FUNCTION_BLOCK PID_GAIN_TRANSITION (* Experimental; offline checks only; native export/runtime pending *)
  (* Standard: 61499-2 *)
  (* Version 0.1, 2026-10-20, Guilherme *)
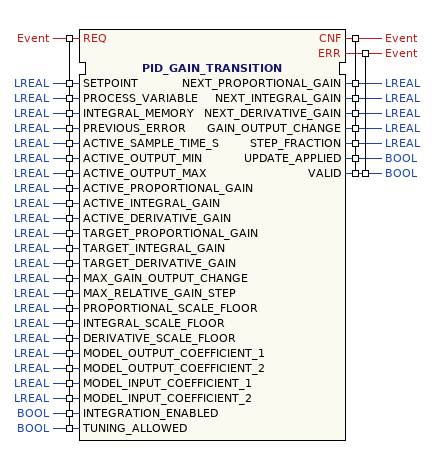
  EVENT_INPUT
    REQ WITH SETPOINT, PROCESS_VARIABLE, INTEGRAL_MEMORY, PREVIOUS_ERROR, ACTIVE_SAMPLE_TIME_S, ACTIVE_OUTPUT_MIN, ACTIVE_OUTPUT_MAX, ACTIVE_PROPORTIONAL_GAIN, ACTIVE_INTEGRAL_GAIN, ACTIVE_DERIVATIVE_GAIN, TARGET_PROPORTIONAL_GAIN, TARGET_INTEGRAL_GAIN, TARGET_DERIVATIVE_GAIN, MAX_GAIN_OUTPUT_CHANGE, MAX_RELATIVE_GAIN_STEP, PROPORTIONAL_SCALE_FLOOR, INTEGRAL_SCALE_FLOOR, DERIVATIVE_SCALE_FLOOR, MODEL_OUTPUT_COEFFICIENT_1, MODEL_OUTPUT_COEFFICIENT_2, MODEL_INPUT_COEFFICIENT_1, MODEL_INPUT_COEFFICIENT_2, INTEGRATION_ENABLED, TUNING_ALLOWED;
  END_EVENT
  EVENT_OUTPUT
    CNF WITH NEXT_PROPORTIONAL_GAIN, NEXT_INTEGRAL_GAIN, NEXT_DERIVATIVE_GAIN, GAIN_OUTPUT_CHANGE, STEP_FRACTION, UPDATE_APPLIED, VALID;
    ERR WITH VALID;
  END_EVENT
  VAR_INPUT
    SETPOINT : LREAL;
    PROCESS_VARIABLE : LREAL;
    INTEGRAL_MEMORY : LREAL;
    PREVIOUS_ERROR : LREAL;
    ACTIVE_SAMPLE_TIME_S : LREAL;
    ACTIVE_OUTPUT_MIN : LREAL;
    ACTIVE_OUTPUT_MAX : LREAL;
    ACTIVE_PROPORTIONAL_GAIN : LREAL;
    ACTIVE_INTEGRAL_GAIN : LREAL;
    ACTIVE_DERIVATIVE_GAIN : LREAL;
    TARGET_PROPORTIONAL_GAIN : LREAL;
    TARGET_INTEGRAL_GAIN : LREAL;
    TARGET_DERIVATIVE_GAIN : LREAL;
    MAX_GAIN_OUTPUT_CHANGE : LREAL;
    MAX_RELATIVE_GAIN_STEP : LREAL;
    PROPORTIONAL_SCALE_FLOOR : LREAL;
    INTEGRAL_SCALE_FLOOR : LREAL;
    DERIVATIVE_SCALE_FLOOR : LREAL;
    MODEL_OUTPUT_COEFFICIENT_1 : LREAL;
    MODEL_OUTPUT_COEFFICIENT_2 : LREAL;
    MODEL_INPUT_COEFFICIENT_1 : LREAL;
    MODEL_INPUT_COEFFICIENT_2 : LREAL;
    INTEGRATION_ENABLED : BOOL;
    TUNING_ALLOWED : BOOL;
  END_VAR
  VAR_OUTPUT
    NEXT_PROPORTIONAL_GAIN : LREAL;
    NEXT_INTEGRAL_GAIN : LREAL;
    NEXT_DERIVATIVE_GAIN : LREAL;
    GAIN_OUTPUT_CHANGE : LREAL;
    STEP_FRACTION : LREAL;
    UPDATE_APPLIED : BOOL;
    VALID : BOOL;
  END_VAR
  VAR
    CURRENT_ERROR : LREAL;
    NEXT_INTEGRAL : LREAL;
    CURRENT_DERIVATIVE : LREAL;
    OLD_RAW : LREAL;
    NEW_RAW : LREAL;
    DELTA_P : LREAL;
    DELTA_I : LREAL;
    DELTA_D : LREAL;
    FULL_EFFECT : LREAL;
    MAGNITUDE : LREAL;
    SCALE : LREAL;
    RELATIVE_STEP : LREAL;
    FRACTION_LIMIT : LREAL;
    CANDIDATE_P : LREAL;
    CANDIDATE_I : LREAL;
    CANDIDATE_D : LREAL;
    Q0 : LREAL;
    Q1 : LREAL;
    Q2 : LREAL;
    A1 : LREAL;
    A2 : LREAL;
    A3 : LREAL;
    A4 : LREAL;
    DENOMINATOR : LREAL;
    B1 : LREAL;
    B2 : LREAL;
    B3 : LREAL;
    C1 : LREAL;
    C2 : LREAL;
    D1 : LREAL;
    CANDIDATE_VALID : BOOL;
  END_VAR
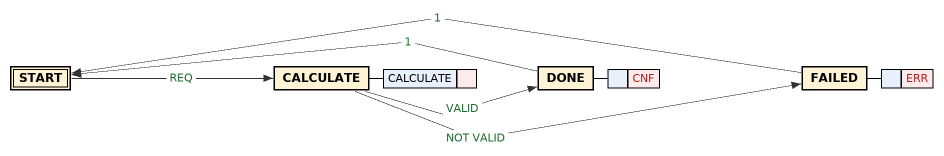
  EC_STATES
    START;
    CALCULATE : CALCULATE;
    DONE : -> CNF;
    FAILED : -> ERR;
  END_STATES
  EC_TRANSITIONS
    START TO CALCULATE := REQ;
    CALCULATE TO DONE := VALID;
    CALCULATE TO FAILED := NOT VALID;
    DONE TO START := 1;
    FAILED TO START := 1;
  END_TRANSITIONS
  ALGORITHM CALCULATE IN ST:
VALID := (SETPOINT >= -1.0E+100) AND (SETPOINT <= 1.0E+100) AND (PROCESS_VARIABLE >= -1.0E+100) AND (PROCESS_VARIABLE <= 1.0E+100) AND (INTEGRAL_MEMORY >= -1.0E+100) AND (INTEGRAL_MEMORY <= 1.0E+100) AND (PREVIOUS_ERROR >= -1.0E+100) AND (PREVIOUS_ERROR <= 1.0E+100) AND (ACTIVE_SAMPLE_TIME_S >= -1.0E+100) AND (ACTIVE_SAMPLE_TIME_S <= 1.0E+100) AND (ACTIVE_OUTPUT_MIN >= -1.0E+100) AND (ACTIVE_OUTPUT_MIN <= 1.0E+100) AND (ACTIVE_OUTPUT_MAX >= -1.0E+100) AND (ACTIVE_OUTPUT_MAX <= 1.0E+100) AND (ACTIVE_PROPORTIONAL_GAIN >= -1.0E+100) AND (ACTIVE_PROPORTIONAL_GAIN <= 1.0E+100) AND (ACTIVE_INTEGRAL_GAIN >= -1.0E+100) AND (ACTIVE_INTEGRAL_GAIN <= 1.0E+100) AND (ACTIVE_DERIVATIVE_GAIN >= -1.0E+100) AND (ACTIVE_DERIVATIVE_GAIN <= 1.0E+100) AND (MAX_GAIN_OUTPUT_CHANGE >= -1.0E+100) AND (MAX_GAIN_OUTPUT_CHANGE <= 1.0E+100) AND (MAX_RELATIVE_GAIN_STEP >= -1.0E+100) AND (MAX_RELATIVE_GAIN_STEP <= 1.0E+100) AND (PROPORTIONAL_SCALE_FLOOR >= -1.0E+100) AND (PROPORTIONAL_SCALE_FLOOR <= 1.0E+100) AND (INTEGRAL_SCALE_FLOOR >= -1.0E+100) AND (INTEGRAL_SCALE_FLOOR <= 1.0E+100) AND (DERIVATIVE_SCALE_FLOOR >= -1.0E+100) AND (DERIVATIVE_SCALE_FLOOR <= 1.0E+100) AND (ACTIVE_SAMPLE_TIME_S > 0.0) AND (ACTIVE_OUTPUT_MIN < ACTIVE_OUTPUT_MAX) AND (MAX_GAIN_OUTPUT_CHANGE > 0.0) AND (MAX_RELATIVE_GAIN_STEP > 0.0) AND (MAX_RELATIVE_GAIN_STEP <= 1.0) AND (PROPORTIONAL_SCALE_FLOOR > 0.0) AND (INTEGRAL_SCALE_FLOOR > 0.0) AND (DERIVATIVE_SCALE_FLOOR > 0.0);
UPDATE_APPLIED := FALSE;
GAIN_OUTPUT_CHANGE := 0.0;
STEP_FRACTION := 0.0;
IF VALID THEN
NEXT_PROPORTIONAL_GAIN := ACTIVE_PROPORTIONAL_GAIN;
NEXT_INTEGRAL_GAIN := ACTIVE_INTEGRAL_GAIN;
NEXT_DERIVATIVE_GAIN := ACTIVE_DERIVATIVE_GAIN;
IF TUNING_ALLOWED AND INTEGRATION_ENABLED THEN
CANDIDATE_VALID := (TARGET_PROPORTIONAL_GAIN >= -1.0E+100) AND (TARGET_PROPORTIONAL_GAIN <= 1.0E+100) AND (TARGET_INTEGRAL_GAIN >= -1.0E+100) AND (TARGET_INTEGRAL_GAIN <= 1.0E+100) AND (TARGET_DERIVATIVE_GAIN >= -1.0E+100) AND (TARGET_DERIVATIVE_GAIN <= 1.0E+100) AND (MODEL_OUTPUT_COEFFICIENT_1 >= -1.0E+100) AND (MODEL_OUTPUT_COEFFICIENT_1 <= 1.0E+100) AND (MODEL_OUTPUT_COEFFICIENT_2 >= -1.0E+100) AND (MODEL_OUTPUT_COEFFICIENT_2 <= 1.0E+100) AND (MODEL_INPUT_COEFFICIENT_1 >= -1.0E+100) AND (MODEL_INPUT_COEFFICIENT_1 <= 1.0E+100) AND (MODEL_INPUT_COEFFICIENT_2 >= -1.0E+100) AND (MODEL_INPUT_COEFFICIENT_2 <= 1.0E+100) AND (TARGET_PROPORTIONAL_GAIN >= 0.0) AND (TARGET_INTEGRAL_GAIN >= 0.0) AND (TARGET_DERIVATIVE_GAIN >= 0.0);
IF CANDIDATE_VALID THEN
CURRENT_ERROR := SETPOINT - PROCESS_VARIABLE;
NEXT_INTEGRAL := INTEGRAL_MEMORY + ACTIVE_SAMPLE_TIME_S / 2.0 * (CURRENT_ERROR + PREVIOUS_ERROR);
CURRENT_DERIVATIVE := (CURRENT_ERROR - PREVIOUS_ERROR) / ACTIVE_SAMPLE_TIME_S;
OLD_RAW := ACTIVE_PROPORTIONAL_GAIN * CURRENT_ERROR + ACTIVE_INTEGRAL_GAIN * NEXT_INTEGRAL + ACTIVE_DERIVATIVE_GAIN * CURRENT_DERIVATIVE;
DELTA_P := TARGET_PROPORTIONAL_GAIN - ACTIVE_PROPORTIONAL_GAIN;
DELTA_I := TARGET_INTEGRAL_GAIN - ACTIVE_INTEGRAL_GAIN;
DELTA_D := TARGET_DERIVATIVE_GAIN - ACTIVE_DERIVATIVE_GAIN;
FULL_EFFECT := DELTA_P * CURRENT_ERROR + DELTA_I * NEXT_INTEGRAL + DELTA_D * CURRENT_DERIVATIVE;
CANDIDATE_VALID := (CURRENT_ERROR >= -1.0E+100) AND (CURRENT_ERROR <= 1.0E+100) AND (NEXT_INTEGRAL >= -1.0E+100) AND (NEXT_INTEGRAL <= 1.0E+100) AND (CURRENT_DERIVATIVE >= -1.0E+100) AND (CURRENT_DERIVATIVE <= 1.0E+100) AND (OLD_RAW >= -1.0E+100) AND (OLD_RAW <= 1.0E+100) AND (FULL_EFFECT >= -1.0E+100) AND (FULL_EFFECT <= 1.0E+100) AND (OLD_RAW >= ACTIVE_OUTPUT_MIN) AND (OLD_RAW <= ACTIVE_OUTPUT_MAX);
IF CANDIDATE_VALID THEN
STEP_FRACTION := 1.0;
MAGNITUDE := FULL_EFFECT;
IF MAGNITUDE < 0.0 THEN
MAGNITUDE := -MAGNITUDE;
END_IF;
IF MAGNITUDE > MAX_GAIN_OUTPUT_CHANGE THEN
STEP_FRACTION := MAX_GAIN_OUTPUT_CHANGE / MAGNITUDE;
END_IF;
SCALE := ACTIVE_PROPORTIONAL_GAIN;
IF SCALE < 0.0 THEN
SCALE := -SCALE;
END_IF;
IF SCALE < PROPORTIONAL_SCALE_FLOOR THEN
SCALE := PROPORTIONAL_SCALE_FLOOR;
END_IF;
MAGNITUDE := DELTA_P;
IF MAGNITUDE < 0.0 THEN
MAGNITUDE := -MAGNITUDE;
END_IF;
RELATIVE_STEP := MAGNITUDE / SCALE;
IF RELATIVE_STEP > MAX_RELATIVE_GAIN_STEP THEN
FRACTION_LIMIT := MAX_RELATIVE_GAIN_STEP / RELATIVE_STEP;
IF FRACTION_LIMIT < STEP_FRACTION THEN
STEP_FRACTION := FRACTION_LIMIT;
END_IF;
END_IF;
CANDIDATE_P := ACTIVE_PROPORTIONAL_GAIN + STEP_FRACTION * DELTA_P;
SCALE := ACTIVE_INTEGRAL_GAIN;
IF SCALE < 0.0 THEN
SCALE := -SCALE;
END_IF;
IF SCALE < INTEGRAL_SCALE_FLOOR THEN
SCALE := INTEGRAL_SCALE_FLOOR;
END_IF;
MAGNITUDE := DELTA_I;
IF MAGNITUDE < 0.0 THEN
MAGNITUDE := -MAGNITUDE;
END_IF;
RELATIVE_STEP := MAGNITUDE / SCALE;
IF RELATIVE_STEP > MAX_RELATIVE_GAIN_STEP THEN
FRACTION_LIMIT := MAX_RELATIVE_GAIN_STEP / RELATIVE_STEP;
IF FRACTION_LIMIT < STEP_FRACTION THEN
STEP_FRACTION := FRACTION_LIMIT;
END_IF;
END_IF;
CANDIDATE_I := ACTIVE_INTEGRAL_GAIN + STEP_FRACTION * DELTA_I;
SCALE := ACTIVE_DERIVATIVE_GAIN;
IF SCALE < 0.0 THEN
SCALE := -SCALE;
END_IF;
IF SCALE < DERIVATIVE_SCALE_FLOOR THEN
SCALE := DERIVATIVE_SCALE_FLOOR;
END_IF;
MAGNITUDE := DELTA_D;
IF MAGNITUDE < 0.0 THEN
MAGNITUDE := -MAGNITUDE;
END_IF;
RELATIVE_STEP := MAGNITUDE / SCALE;
IF RELATIVE_STEP > MAX_RELATIVE_GAIN_STEP THEN
FRACTION_LIMIT := MAX_RELATIVE_GAIN_STEP / RELATIVE_STEP;
IF FRACTION_LIMIT < STEP_FRACTION THEN
STEP_FRACTION := FRACTION_LIMIT;
END_IF;
END_IF;
CANDIDATE_D := ACTIVE_DERIVATIVE_GAIN + STEP_FRACTION * DELTA_D;
CANDIDATE_P := ACTIVE_PROPORTIONAL_GAIN + STEP_FRACTION * DELTA_P;
CANDIDATE_I := ACTIVE_INTEGRAL_GAIN + STEP_FRACTION * DELTA_I;
CANDIDATE_D := ACTIVE_DERIVATIVE_GAIN + STEP_FRACTION * DELTA_D;
NEW_RAW := CANDIDATE_P * CURRENT_ERROR + CANDIDATE_I * NEXT_INTEGRAL + CANDIDATE_D * CURRENT_DERIVATIVE;
Q0 := CANDIDATE_P + CANDIDATE_I * ACTIVE_SAMPLE_TIME_S / 2.0 + CANDIDATE_D / ACTIVE_SAMPLE_TIME_S;
Q1 := -CANDIDATE_P + CANDIDATE_I * ACTIVE_SAMPLE_TIME_S / 2.0 - 2.0 * CANDIDATE_D / ACTIVE_SAMPLE_TIME_S;
Q2 := CANDIDATE_D / ACTIVE_SAMPLE_TIME_S;
A1 := -1.0 - MODEL_OUTPUT_COEFFICIENT_1 + MODEL_INPUT_COEFFICIENT_1 * Q0;
A2 := MODEL_OUTPUT_COEFFICIENT_1 - MODEL_OUTPUT_COEFFICIENT_2 + MODEL_INPUT_COEFFICIENT_1 * Q1 + MODEL_INPUT_COEFFICIENT_2 * Q0;
A3 := MODEL_OUTPUT_COEFFICIENT_2 + MODEL_INPUT_COEFFICIENT_1 * Q2 + MODEL_INPUT_COEFFICIENT_2 * Q1;
A4 := MODEL_INPUT_COEFFICIENT_2 * Q2;
CANDIDATE_VALID := (CANDIDATE_P >= -1.0E+100) AND (CANDIDATE_P <= 1.0E+100) AND (CANDIDATE_I >= -1.0E+100) AND (CANDIDATE_I <= 1.0E+100) AND (CANDIDATE_D >= -1.0E+100) AND (CANDIDATE_D <= 1.0E+100) AND (NEW_RAW >= -1.0E+100) AND (NEW_RAW <= 1.0E+100) AND (A1 >= -1.0E+100) AND (A1 <= 1.0E+100) AND (A2 >= -1.0E+100) AND (A2 <= 1.0E+100) AND (A3 >= -1.0E+100) AND (A3 <= 1.0E+100) AND (A4 >= -1.0E+100) AND (A4 <= 1.0E+100) AND (NEW_RAW >= ACTIVE_OUTPUT_MIN) AND (NEW_RAW <= ACTIVE_OUTPUT_MAX);
IF CANDIDATE_VALID THEN
CANDIDATE_VALID := (A4 > -1.0) AND (A4 < 1.0);
IF CANDIDATE_VALID THEN
DENOMINATOR := 1.0 - A4 * A4;
CANDIDATE_VALID := DENOMINATOR > 1.0E-12;
IF CANDIDATE_VALID THEN
B1 := (A1 - A4 * A3) / DENOMINATOR;
B2 := (A2 - A4 * A2) / DENOMINATOR;
B3 := (A3 - A4 * A1) / DENOMINATOR;
CANDIDATE_VALID := (B1 >= -1.0E+100) AND (B1 <= 1.0E+100) AND (B2 >= -1.0E+100) AND (B2 <= 1.0E+100) AND (B3 >= -1.0E+100) AND (B3 <= 1.0E+100);
END_IF;
END_IF;
END_IF;
IF CANDIDATE_VALID THEN
CANDIDATE_VALID := (B3 > -1.0) AND (B3 < 1.0);
IF CANDIDATE_VALID THEN
DENOMINATOR := 1.0 - B3 * B3;
CANDIDATE_VALID := DENOMINATOR > 1.0E-12;
IF CANDIDATE_VALID THEN
C1 := (B1 - B3 * B2) / DENOMINATOR;
C2 := (B2 - B3 * B1) / DENOMINATOR;
CANDIDATE_VALID := (C1 >= -1.0E+100) AND (C1 <= 1.0E+100) AND (C2 >= -1.0E+100) AND (C2 <= 1.0E+100);
END_IF;
END_IF;
END_IF;
IF CANDIDATE_VALID THEN
CANDIDATE_VALID := (C2 > -1.0) AND (C2 < 1.0);
IF CANDIDATE_VALID THEN
DENOMINATOR := 1.0 - C2 * C2;
CANDIDATE_VALID := DENOMINATOR > 1.0E-12;
IF CANDIDATE_VALID THEN
D1 := (C1 - C2 * C1) / DENOMINATOR;
CANDIDATE_VALID := (D1 >= -1.0E+100) AND (D1 <= 1.0E+100);
END_IF;
END_IF;
END_IF;
IF CANDIDATE_VALID THEN
CANDIDATE_VALID := (D1 > -1.0) AND (D1 < 1.0);
END_IF;
IF CANDIDATE_VALID THEN
NEXT_PROPORTIONAL_GAIN := CANDIDATE_P;
NEXT_INTEGRAL_GAIN := CANDIDATE_I;
NEXT_DERIVATIVE_GAIN := CANDIDATE_D;
GAIN_OUTPUT_CHANGE := NEW_RAW - OLD_RAW;
UPDATE_APPLIED := (DELTA_P <> 0.0) OR (DELTA_I <> 0.0) OR (DELTA_D <> 0.0);
END_IF;
IF NOT CANDIDATE_VALID THEN
STEP_FRACTION := 0.0;
END_IF;
END_IF;
END_IF;
END_IF;
END_IF;
  END_ALGORITHM
END_FUNCTION_BLOCK
